(* IEC 61131-3 sources: plcassist-cli/packages/volt-lsp-iec/test-corpus/pro2193/Device/Plc Logic/Application/09 Misc/Library Manager/CAA NetBaseSrv, 33 files *)

(* ---- ASYNCGLOB.gvl ---- *)
VAR_GLOBAL
	G_XGLOBALLIBINITDONE : BOOL := AsyncInitTask();
	GC_STASKRW : STRING := 'CAA_NetBaseServices_RW';
	GC_STASKOPENER : STRING := gc_sTaskRW;
END_VAR

(* ---- CAA_ASM_CONSTANTS.gvl ---- *)
VAR_GLOBAL
	UDP_PEER_OPEN_JOB_ID : UDINT := 16#50001;
	UDP_PEER_CLOSE_JOB_ID : UDINT := 16#50002;
	UDP_RECEIVE_JOB_ID : UDINT := 16#50003;
	UDP_SEND_JOB_ID : UDINT := 16#50004;
	TCP_SERVER_OPEN_JOB_ID : UDINT := 16#50005;
	TCP_CLIENT_OPEN_JOB_ID : UDINT := 16#50006;
	TCP_CONNECTION_OPEN_JOB_ID : UDINT := 16#50007;
	TCP_CLOSE_JOB_ID : UDINT := 16#50008;
	TCP_READ_JOB_ID : UDINT := 16#50009;
	TCP_WRITE_JOB_ID : UDINT := 16#5000A;
END_VAR

(* ---- CONSTANTS.gvl ---- *)
VAR_GLOBAL
	GC_FIRST_MULTICAST_IP : UDINT := 16#E0000000;
	GC_LAST_MULTICAST_IP : UDINT := 16#EFFFFFFF;
END_VAR

(* ---- FUNCTIONALITIES.gvl ---- *)
VAR_GLOBAL
	GC_XSUPPORTSTCPCLIENTSETADAPTER : BOOL;
END_VAR

(* ---- HOTO.gvl ---- *)
VAR_GLOBAL
	IDUMMY : INT;
END_VAR

(* ---- PARAM.gvl ---- *)
VAR_GLOBAL
	GC_UDITASKRWPRIORITY : UDINT := 240;
	GC_UDITASKOPENERPRIORITY : UDINT := gc_udiTaskRWPriority;
END_VAR

(* ---- VARIABLES.gvl ---- *)
VAR_GLOBAL
	G_HSOCKETCLASS : CAA.HANDLE;
END_VAR

(* ---- VERSIONCONSTANTS.gvl ---- *)
VAR_GLOBAL
	GC_BYVERSION : BYTE := 1;
	GC_BYVERSION_1 : BYTE := 0;
END_VAR

(* ---- ITCPCONNECTION.itf ---- *)
INTERFACE ITCPCONNECTION
END_INTERFACE

METHOD PRVCLOSE : ERROR
VAR_INPUT
	XDUMMY : BOOL;
END_VAR
END_METHOD

METHOD PRVESTABLISH : ERROR
END_METHOD

(* ---- ITCPSERVER.itf ---- *)
INTERFACE ITCPSERVER
END_INTERFACE

METHOD PRVADDCONNECTION : ERROR
VAR_INPUT
	CONNECTION : ITCPConnection;
END_VAR
END_METHOD

METHOD PRVREMOVECONNECTION : ERROR
VAR_INPUT
	CONNECTION : ITCPConnection;
END_VAR
END_METHOD

(* ---- ASYNCINITTASK.fun ---- *)
FUNCTION ASYNCINITTASK : BOOL
END_FUNCTION

(* ---- ASYNCINITTASK2INIT.fun ---- *)
FUNCTION ASYNCINITTASK2INIT : RTS_IEC_RESULT
VAR_INPUT
	PPARAM : __XWORD;
END_VAR
END_FUNCTION

(* ---- DUMMYJOB.fun ---- *)
FUNCTION DUMMYJOB : RTS_IEC_RESULT
VAR_INPUT
	PPARAM : __XWORD;
END_VAR
END_FUNCTION

(* ---- GETSUPPLIERVERSION.fun ---- *)
FUNCTION GETSUPPLIERVERSION : WORD
END_FUNCTION

(* ---- GETTCPSOCKETHANDLE.fun ---- *)
FUNCTION GETTCPSOCKETHANDLE : SysTypes.RTS_IEC_HANDLE
VAR_INPUT
	HCONNECTION : CAA.HANDLE;
END_VAR
END_FUNCTION

(* ---- GETUDPSOCKETHANDLE.fun ---- *)
FUNCTION GETUDPSOCKETHANDLE : SysTypes.RTS_IEC_HANDLE
VAR_INPUT
	HPEER : CAA.HANDLE;
END_VAR
END_FUNCTION

(* ---- IPSTRING_TO_UDINT.fun ---- *)
FUNCTION IPSTRING_TO_UDINT : UDINT
VAR_INPUT
	SIPADDRESS : STRING;
END_VAR
END_FUNCTION

(* ---- IS_MULTICAST_GROUP.fun ---- *)
FUNCTION IS_MULTICAST_GROUP : BOOL
VAR_INPUT
	UDIIPADDRESS : UDINT;
END_VAR
END_FUNCTION

(* ---- UDINT_TO_IPSTRING.fun ---- *)
FUNCTION UDINT_TO_IPSTRING : STRING
VAR_INPUT
	UDIIPADDRESS : UDINT;
END_VAR
END_FUNCTION

(* ---- UDP_GETDATASIZE.fun ---- *)
FUNCTION UDP_GETDATASIZE : CAA.SIZE
VAR_INPUT
	HPEER : CAA.HANDLE;
	PEERROR : POINTER TO ERROR;
END_VAR
END_FUNCTION

(* ---- TCP_CLIENT.fb ---- *)
FUNCTION_BLOCK TCP_CLIENT EXTENDS LTrig
VAR_INPUT
	UDITIMEOUT : UDINT := 0;
	IPADDR : IP_ADDR;
	UIPORT : UINT;
END_VAR
VAR_OUTPUT
	EERROR : ERROR;
	XACTIVE : BOOL;
	HCONNECTION : CAA.HANDLE;
END_VAR
VAR
	_UIPORT : UINT;
	_IPADDR : IP_ADDR;
	_ITFCONNECTION : TCPConnection;
	_TKSTART : CAA.TICK;
	_TCPCONNECTOR : TCP.Connector;
	_REBUILDDETECTRISINGEDGE : BOOL := FALSE;
	_ASYNC : ST_ASYNC;
	_ASYNCCLOSER : ST_ASYNC;
	_ASYNCRESETOUTPUTS : ST_ASYNC;
	_DBHOLDVALVS1TICK : BOOL;
	_DB_XDONE : BOOL;
	_DB_XBUSY : BOOL;
	_DB_XERROR : BOOL;
	_DB_IERROR : INT;
	_DB_EERROR : ERROR;
	_DB_XACTIVE : BOOL;
	_DB_HCONNECTION : CAA.HANDLE;
END_VAR
END_FUNCTION_BLOCK

METHOD FB_EXIT : BOOL
VAR_INPUT
	BINCOPYCODE : BOOL;
END_VAR
END_METHOD

METHOD FB_INIT : BOOL
VAR_INPUT
	BINITRETAINS : BOOL;
	BINCOPYCODE : BOOL;
END_VAR
END_METHOD

METHOD SETADAPTER : ERROR
VAR_INPUT
	IPADDR : IP_ADDR;
END_VAR
END_METHOD

METHOD PRVABORT : BOOL
END_METHOD

METHOD PRVASYNCABORT : RTS_IEC_RESULT
VAR_INPUT
	PPARAM : __XWORD;
END_VAR
END_METHOD

METHOD PRVASYNCCYCLICACTION : RTS_IEC_RESULT
VAR_INPUT
	PPARAM : __XWORD;
END_VAR
END_METHOD

METHOD PRVASYNCRESETOUTPUTS : RTS_IEC_RESULT
VAR_INPUT
	PPARAM : __XWORD;
END_VAR
END_METHOD

METHOD PRVCLOSE : BOOL
END_METHOD

METHOD PRVCYCLICACTION : BOOL
END_METHOD

METHOD PRVRESETOUTPUTS : BOOL
END_METHOD

METHOD PRVSTART : BOOL
END_METHOD

(* ---- TCP_CONNECTION.fb ---- *)
FUNCTION_BLOCK TCP_CONNECTION EXTENDS LTrig
VAR_INPUT
	HSERVER : CAA.HANDLE;
END_VAR
VAR_OUTPUT
	EERROR : ERROR;
	XACTIVE : BOOL;
	HCONNECTION : CAA.HANDLE;
END_VAR
VAR
	HCONNECTIONTMP : CAA.HANDLE;
	ITFSERVER : ITCPServer;
	PSERVER : POINTER TO TCP_Server;
	IINPUTERROR : ERROR;
	ITFCONNECTION : TCPConnection;
	_ASYNC : ST_ASYNC;
	_ASYNCCLOSER : ST_ASYNC;
	_ASYNCRESETOUTPUTS : ST_ASYNC;
	_REBUILDDETECTRISINGEDGE : BOOL := FALSE;
	_DBHOLDVALVS1TICK : BOOL;
	_DB_XDONE : BOOL;
	_DB_XBUSY : BOOL;
	_DB_XERROR : BOOL;
	_DB_IERROR : INT;
	_DB_EERROR : ERROR;
	_DB_XACTIVE : BOOL;
	_DB_HCONNECTION : CAA.HANDLE;
	IPADDRESS : SysSocket.INADDR;
END_VAR
END_FUNCTION_BLOCK

METHOD FB_EXIT : BOOL
VAR_INPUT
	BINCOPYCODE : BOOL;
END_VAR
END_METHOD

METHOD FB_INIT : BOOL
VAR_INPUT
	BINITRETAINS : BOOL;
	BINCOPYCODE : BOOL;
END_VAR
END_METHOD

METHOD PRVABORT : BOOL
END_METHOD

METHOD PRVASYNCABORT : RTS_IEC_RESULT
VAR_INPUT
	PPARAM : __XWORD;
END_VAR
END_METHOD

METHOD PRVASYNCCYCLICACTION : RTS_IEC_RESULT
VAR_INPUT
	PPARAM : __XWORD;
END_VAR
END_METHOD

METHOD PRVASYNCRESETOUTPUTS : RTS_IEC_RESULT
VAR_INPUT
	PPARAM : __XWORD;
END_VAR
END_METHOD

METHOD PRVCLOSE : BOOL
END_METHOD

METHOD PRVCYCLICACTION : BOOL
END_METHOD

METHOD PRVRESETOUTPUTS : BOOL
END_METHOD

METHOD PRVSTART : BOOL
END_METHOD

(* ---- TCP_READ.fb ---- *)
FUNCTION_BLOCK TCP_READ EXTENDS LTrig
VAR_INPUT
	HCONNECTION : CAA.HANDLE;
	SZSIZE : CAA.SIZE;
	PDATA : CAA.PVOID;
END_VAR
VAR_OUTPUT
	EERROR : ERROR;
	XREADY : BOOL;
	SZCOUNT : CAA.SIZE;
END_VAR
VAR
	IINPUTERROR : ERROR;
	ITFCONNECTION : ITCPConnection;
	_ASYNC : ST_ASYNC;
	_DBHOLDVALVS1TICK : BOOL;
	_DB_XDONE : BOOL;
	_DB_XBUSY : BOOL;
	_DB_XERROR : BOOL;
	_DB_IERROR : INT;
	_DB_EERROR : ERROR;
	_DB_XREADY : BOOL;
	_DB_SZCOUNT : CAA.SIZE;
END_VAR
END_FUNCTION_BLOCK

METHOD FB_EXIT : BOOL
VAR_INPUT
	BINCOPYCODE : BOOL;
END_VAR
END_METHOD

METHOD FB_INIT : BOOL
VAR_INPUT
	BINITRETAINS : BOOL;
	BINCOPYCODE : BOOL;
END_VAR
END_METHOD

METHOD PRVABORT : BOOL
END_METHOD

METHOD PRVASYNCCYCLICACTION : RTS_IEC_RESULT
VAR_INPUT
	PPARAM : __XWORD;
END_VAR
END_METHOD

METHOD PRVCYCLICACTION : BOOL
END_METHOD

METHOD PRVRESETOUTPUTS : BOOL
END_METHOD

METHOD PRVSTART : BOOL
END_METHOD

(* ---- TCP_READBUFFER.fb ---- *)
FUNCTION_BLOCK TCP_READBUFFER EXTENDS LTrig
VAR_INPUT
	HCONNECTION : CAA.HANDLE;
END_VAR
VAR_OUTPUT
	EERROR : ERROR;
	XREADY : BOOL;
	HBUFFER : CAA.HANDLE;
END_VAR
VAR
	IINPUTERROR : ERROR;
	ITFCONNECTION : ITCPConnection;
	_ASYNC : ST_ASYNC;
	_DBHOLDVALVS1TICK : BOOL;
	_DB_XDONE : BOOL;
	_DB_XBUSY : BOOL;
	_DB_XERROR : BOOL;
	_DB_IERROR : INT;
	_DB_EERROR : ERROR;
	_DB_XREADY : BOOL;
	_DB_HBUFFER : CAA.HANDLE;
END_VAR
END_FUNCTION_BLOCK

METHOD FB_EXIT : BOOL
VAR_INPUT
	BINCOPYCODE : BOOL;
END_VAR
END_METHOD

METHOD FB_INIT : BOOL
VAR_INPUT
	BINITRETAINS : BOOL;
	BINCOPYCODE : BOOL;
END_VAR
END_METHOD

METHOD PRVABORT : BOOL
END_METHOD

METHOD PRVASYNCCYCLICACTION : RTS_IEC_RESULT
VAR_INPUT
	PPARAM : __XWORD;
END_VAR
END_METHOD

METHOD PRVCYCLICACTION : BOOL
END_METHOD

METHOD PRVRESETOUTPUTS : BOOL
END_METHOD

METHOD PRVSTART : BOOL
END_METHOD

(* ---- TCP_SERVER.fb ---- *)
FUNCTION_BLOCK TCP_SERVER EXTENDS LTrig
VAR_INPUT
	IPADDR : IP_ADDR := STRUCT(sAddr := '0.0.0.0');
	UIPORT : UINT;
END_VAR
VAR_OUTPUT
	EERROR : ERROR;
	HSERVER : CAA.HANDLE;
END_VAR
VAR
	_UIPORT : UINT;
	_IPADDR : IP_ADDR;
	_LSTCONNECTIONS : LAT.List;
	_ITFSERVER : ITCPServer;
	_PSERVER : POINTER TO TCP_Server;
	_TCPLISTENER : TCP.Listener;
	_ESTATE : SERVER_STATE := SERVER_STATE.NOT_LISTENING;
	_REBUILDDETECTRISINGEDGE : BOOL := FALSE;
	_ASYNC : ST_ASYNC;
	_ASYNCCLOSER : ST_ASYNC;
	_ASYNCRESETOUTPUTS : ST_ASYNC;
	_DBHOLDVALVS1TICK : BOOL;
	_DB_XDONE : BOOL;
	_DB_XBUSY : BOOL;
	_DB_XERROR : BOOL;
	_DB_IERROR : INT;
	_DB_EERROR : ERROR;
	_DB_HSERVER : CAA.HANDLE;
END_VAR
END_FUNCTION_BLOCK

METHOD FB_EXIT : BOOL
VAR_INPUT
	BINCOPYCODE : BOOL;
END_VAR
END_METHOD

METHOD FB_INIT : BOOL
VAR_INPUT
	BINITRETAINS : BOOL;
	BINCOPYCODE : BOOL;
END_VAR
END_METHOD

METHOD PRVABORT : BOOL
END_METHOD

METHOD PRVADDCONNECTION : ERROR
VAR_INPUT
	CONNECTION : ITCPConnection;
END_VAR
END_METHOD

METHOD PRVASYNCABORT : RTS_IEC_RESULT
VAR_INPUT
	PPARAM : __XWORD;
END_VAR
END_METHOD

METHOD PRVASYNCCYCLICACTION : RTS_IEC_RESULT
VAR_INPUT
	PPARAM : __XWORD;
END_VAR
END_METHOD

METHOD PRVASYNCRESETOUTPUTS : RTS_IEC_RESULT
VAR_INPUT
	PPARAM : __XWORD;
END_VAR
END_METHOD

METHOD PRVCLOSE
END_METHOD

METHOD PRVCYCLICACTION : BOOL
END_METHOD

METHOD PRVREMOVECONNECTION : ERROR
VAR_INPUT
	CONNECTION : ITCPConnection;
END_VAR
END_METHOD

METHOD PRVRESETOUTPUTS : BOOL
END_METHOD

METHOD PRVSTART : BOOL
END_METHOD

(* ---- TCP_WRITE.fb ---- *)
FUNCTION_BLOCK TCP_WRITE EXTENDS ETrigTo
VAR_INPUT
	HCONNECTION : CAA.HANDLE;
	SZSIZE : CAA.SIZE;
	PDATA : CAA.PVOID;
END_VAR
VAR_OUTPUT
	EERROR : ERROR;
END_VAR
VAR
	ESEGBUFMANERROR : SBM.ERROR;
	IINPUTERROR : ERROR;
	ITFCONNECTION : ITCPConnection;
	_SZSENTBYTES : CAA.SIZE;
	_EWRITESTATE : TCP_WRITE_STATE;
	_ASYNC : ST_ASYNC;
	_ASYNCCLOSER : ST_ASYNC;
	_ASYNCRESETOUTPUTS : ST_ASYNC;
	_DBHOLDVALVS1TICK : BOOL;
	_DB_XDONE : BOOL;
	_DB_XBUSY : BOOL;
	_DB_XERROR : BOOL;
	_DB_IERROR : INT;
	_DB_EERROR : ERROR;
END_VAR
END_FUNCTION_BLOCK

METHOD FB_EXIT : BOOL
VAR_INPUT
	BINCOPYCODE : BOOL;
END_VAR
END_METHOD

METHOD FB_INIT : BOOL
VAR_INPUT
	BINITRETAINS : BOOL;
	BINCOPYCODE : BOOL;
END_VAR
END_METHOD

METHOD PRVABORT : BOOL
END_METHOD

METHOD PRVASYNCABORT : RTS_IEC_RESULT
VAR_INPUT
	PPARAM : __XWORD;
END_VAR
END_METHOD

METHOD PRVASYNCCYCLICACTION : RTS_IEC_RESULT
VAR_INPUT
	PPARAM : __XWORD;
END_VAR
END_METHOD

METHOD PRVCYCLICACTION : BOOL
END_METHOD

METHOD PRVRESETOUTPUTS : BOOL
END_METHOD

METHOD PRVSTART : BOOL
END_METHOD

(* ---- TCP_WRITEBUFFER.fb ---- *)
FUNCTION_BLOCK TCP_WRITEBUFFER EXTENDS ETrigTo
VAR_INPUT
	HCONNECTION : CAA.HANDLE;
	HBUFFER : CAA.HANDLE;
END_VAR
VAR_OUTPUT
	EERROR : ERROR;
END_VAR
VAR
	_HBUFFER : CAA.HANDLE;
	IINPUTERROR : ERROR;
	ITFCONNECTION : ITCPConnection;
	_SZSENTBYTES : CAA.SIZE;
	_EWRITESTATE : TCP_WRITE_STATE;
	_ASYNC : ST_ASYNC;
	_ASYNCCLOSER : ST_ASYNC;
	_ASYNCRESETOUTPUTS : ST_ASYNC;
	_DBHOLDVALVS1TICK : BOOL;
	_DB_XDONE : BOOL;
	_DB_XBUSY : BOOL;
	_DB_XERROR : BOOL;
	_DB_IERROR : INT;
	_DB_EERROR : ERROR;
END_VAR
END_FUNCTION_BLOCK

METHOD FB_EXIT : BOOL
VAR_INPUT
	BINCOPYCODE : BOOL;
END_VAR
END_METHOD

METHOD FB_INIT : BOOL
VAR_INPUT
	BINITRETAINS : BOOL;
	BINCOPYCODE : BOOL;
END_VAR
END_METHOD

METHOD PRVABORT : BOOL
END_METHOD

METHOD PRVASYNCABORT : RTS_IEC_RESULT
VAR_INPUT
	PPARAM : __XWORD;
END_VAR
END_METHOD

METHOD PRVASYNCCYCLICACTION : RTS_IEC_RESULT
VAR_INPUT
	PPARAM : __XWORD;
END_VAR
END_METHOD

METHOD PRVASYNCRESETOUTPUTS : RTS_IEC_RESULT
VAR_INPUT
	PPARAM : __XWORD;
END_VAR
END_METHOD

METHOD PRVCYCLICACTION : BOOL
END_METHOD

METHOD PRVRESETOUTPUTS : BOOL
END_METHOD

METHOD PRVSTART : BOOL
END_METHOD

(* ---- TCPCONNECTION.fb ---- *)
FUNCTION_BLOCK TCPCONNECTION EXTENDS Element
VAR
	TCPSTREAM : TCP.Stream;
	HSOCKET : SysTypes.RTS_IEC_HANDLE := SysTypes.RTS_INVALID_HANDLE;
	ESTATE : CONNECTION_STATE := CONNECTION_STATE.LISTEN;
	_PUSHBACK1READBYTE_DATA : BYTE;
	_PUSHBACK1READBYTE_CALLED : BOOL;
	PRVSOCKETHANDLE : RTS_IEC_HANDLE;
	PRVSTATE : CONNECTION_STATE;
	PRVSTREAM : POINTER TO TCP.Stream;
END_VAR
END_FUNCTION_BLOCK

METHOD FB_EXIT : BOOL
VAR_INPUT
	BINCOPYCODE : BOOL;
END_VAR
END_METHOD

METHOD SETPUSHBACK1READBYTE
VAR_INPUT
	DATA : BYTE;
	CALLED : BOOL;
END_VAR
END_METHOD

METHOD PRVCLOSE : ERROR
VAR_INPUT
	XDUMMY : BOOL;
END_VAR
END_METHOD

METHOD PRVESTABLISH : ERROR
END_METHOD

(* ---- UDP_PEER.fb ---- *)
FUNCTION_BLOCK UDP_PEER EXTENDS LTrig
VAR_INPUT
	IPADDR : IP_ADDR := STRUCT(sAddr := '0.0.0.0');
	UIPORT : UINT;
	IPMULTICAST : IP_ADDR := STRUCT(sAddr := '255.255.255.255');
END_VAR
VAR_OUTPUT
	EERROR : ERROR;
	XACTIVE : BOOL;
	HPEER : CAA.HANDLE;
END_VAR
VAR
	_UDIIPADDRESS : UDINT;
	_UDIMCIPADDRESS : UDINT;
	_UDPDRIVER : UDP.UDPDriver;
	_UDPPORT : UDP.Port;
END_VAR
END_FUNCTION_BLOCK

METHOD FB_EXIT : BOOL
VAR_INPUT
	BINCOPYCODE : BOOL;
END_VAR
END_METHOD

METHOD PRVABORT : BOOL
END_METHOD

METHOD PRVCLOSE
END_METHOD

METHOD PRVCYCLICACTION : BOOL
END_METHOD

METHOD PRVRESETOUTPUTS : BOOL
END_METHOD

METHOD PRVSTART : BOOL
END_METHOD

(* ---- UDP_RECEIVE.fb ---- *)
FUNCTION_BLOCK UDP_RECEIVE EXTENDS LTrig
VAR_INPUT
	HPEER : CAA.HANDLE;
	SZSIZE : CAA.SIZE;
	PDATA : CAA.PVOID;
END_VAR
VAR_OUTPUT
	EERROR : ERROR;
	XREADY : BOOL;
	IPFROM : IP_ADDR;
	UIPORTFROM : UINT;
	SZCOUNT : CAA.SIZE;
END_VAR
VAR
	_PUDPPORT : POINTER TO UDP.Port;
	IINPUTERROR : ERROR;
END_VAR
END_FUNCTION_BLOCK

METHOD PRVABORT : BOOL
END_METHOD

METHOD PRVCYCLICACTION : BOOL
END_METHOD

METHOD PRVRESETOUTPUTS : BOOL
END_METHOD

METHOD PRVSTART : BOOL
END_METHOD

(* ---- UDP_RECEIVEBUFFER.fb ---- *)
FUNCTION_BLOCK UDP_RECEIVEBUFFER EXTENDS LTrig
VAR_INPUT
	HPEER : CAA.HANDLE;
END_VAR
VAR_OUTPUT
	EERROR : ERROR;
	XREADY : BOOL;
	IPFROM : IP_ADDR;
	UIPORTFROM : UINT;
	HBUFFER : CAA.HANDLE;
END_VAR
VAR
	_PUDPPORT : POINTER TO UDP.Port;
	IINPUTERROR : ERROR;
END_VAR
END_FUNCTION_BLOCK

METHOD PRVABORT : BOOL
END_METHOD

METHOD PRVCYCLICACTION : BOOL
END_METHOD

METHOD PRVRESETOUTPUTS : BOOL
END_METHOD

METHOD PRVSTART : BOOL
END_METHOD

(* ---- UDP_SEND.fb ---- *)
FUNCTION_BLOCK UDP_SEND EXTENDS ETrigTo
VAR_INPUT
	HPEER : CAA.HANDLE;
	IPADDR : IP_ADDR;
	UIPORT : UINT;
	SZSIZE : CAA.SIZE;
	PDATA : CAA.PVOID;
END_VAR
VAR_OUTPUT
	EERROR : ERROR;
END_VAR
VAR
	IINPUTERROR : ERROR;
	_PUDPPORT : POINTER TO UDP.Port;
END_VAR
END_FUNCTION_BLOCK

METHOD PRVABORT : BOOL
END_METHOD

METHOD PRVCYCLICACTION : BOOL
END_METHOD

METHOD PRVRESETOUTPUTS : BOOL
END_METHOD

METHOD PRVSTART : BOOL
END_METHOD

(* ---- UDP_SENDBUFFER.fb ---- *)
FUNCTION_BLOCK UDP_SENDBUFFER EXTENDS ETrigTo
VAR_INPUT
	HPEER : CAA.HANDLE;
	IPADDR : IP_ADDR;
	UIPORT : UINT;
	HBUFFER : CAA.HANDLE;
END_VAR
VAR_OUTPUT
	EERROR : ERROR;
END_VAR
VAR
	_HBUFFER : CAA.HANDLE;
	IINPUTERROR : ERROR;
	_PUDPPORT : POINTER TO UDP.Port;
END_VAR
END_FUNCTION_BLOCK

METHOD FB_EXIT : BOOL
VAR_INPUT
	BINCOPYCODE : BOOL;
END_VAR
END_METHOD

METHOD PRVABORT : BOOL
END_METHOD

METHOD PRVCYCLICACTION : BOOL
END_METHOD

METHOD PRVRESETOUTPUTS : BOOL
END_METHOD

METHOD PRVSTART : BOOL
END_METHOD
